Fanuc KAREL source: KT00816.KL

PROGRAM KT00816
%NOLOCKGROUP
VAR
  B1: BOOLEAN
  B2: BOOLEAN
  OUT: INTEGER
BEGIN
  B1 = TRUE
  B2 = FALSE
  B1 = TRUE
  B2 = FALSE
  OUT = LN(B1)
END KT00816
